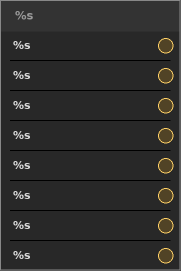
VISUALIZATION FRM_8BitPairDisplay  // 181x271
VAR_IN_OUT
    bBit0_1: BOOL;
    bBit1_1: BOOL;
    bBit2_1: BOOL;
    bBit3_1: BOOL;
    bBit4_1: BOOL;
    bBit5_1: BOOL;
    bBit6_1: BOOL;
    bBit7_1: BOOL;
    
    bBit0_2: BOOL;
    bBit1_2: BOOL;
    bBit2_2: BOOL;
    bBit3_2: BOOL;
    bBit4_2: BOOL;
    bBit5_2: BOOL;
    bBit6_2: BOOL;
    bBit7_2: BOOL;
END_VAR
VAR_INPUT
    sName: STRING;	

    sBitPair0: STRING;
    sBitPair1: STRING;
    sBitPair2: STRING;
    sBitPair3: STRING;
    sBitPair4: STRING;
    sBitPair5: STRING;
    sBitPair6: STRING;
    sBitPair7: STRING;	
END_VAR
    Rectangle (0,30 181x241)
    Textfield (10,40 141x11), "%s", text variable: sBitPair0
    Textfield (10,70 141x11), "%s", text variable: sBitPair1
    Textfield (10,100 141x11), "%s", text variable: sBitPair2
    Textfield (10,130 141x11), "%s", text variable: sBitPair3
    Textfield (10,160 141x11), "%s", text variable: sBitPair4
    Textfield (10,190 151x11), "%s", text variable: sBitPair5
    Textfield (10,220 141x11), "%s", text variable: sBitPair6
    Textfield (10,250 141x11), "%s", text variable: sBitPair7
    Line (10,60) (170,60)
    Line (10,90) (170,90)
    Line (10,120) (170,120)
    Line (10,150) (170,150)
    Line (10,180) (170,180)
    Line (10,210) (170,210)
    Line (10,240) (170,240)
    Textfield (0,0 181x31), "%s", text variable: sName
    Ellipse (158,38 15x15), colour toggle: bBit0_1 AND bBit0_2
    Ellipse (158,68 15x15), colour toggle: bBit1_1 AND bBit1_2
    Ellipse (158,98 15x15), colour toggle: bBit2_1 AND bBit2_2
    Ellipse (158,128 15x15), colour toggle: bBit3_1 AND bBit3_2
    Ellipse (158,158 15x15), colour toggle: bBit4_1 AND bBit4_2
    Ellipse (158,188 15x15), colour toggle: bBit5_1 AND bBit5_2
    Ellipse (158,218 15x15), colour toggle: bBit6_1 AND bBit6_2
    Ellipse (158,248 15x15), colour toggle: bBit7_1 AND bBit7_2
    Ellipse (158,38 15x15), invisible if: NOT (bBit0_1 XOR bBit0_2)
    Ellipse (158,68 15x15), invisible if: NOT (bBit1_1 XOR bBit1_2)
    Ellipse (158,98 15x15), invisible if: NOT (bBit2_1 XOR bBit2_2)
    Ellipse (158,128 15x15), invisible if: NOT (bBit3_1 XOR bBit3_2)
    Ellipse (158,158 15x15), invisible if: NOT (bBit4_1 XOR bBit4_2)
    Ellipse (158,188 15x15), invisible if: NOT (bBit5_1 XOR bBit5_2)
    Ellipse (158,218 15x15), invisible if: NOT (bBit6_1 XOR bBit6_2)
    Ellipse (158,248 15x15), invisible if: NOT (bBit7_1 XOR bBit7_2)
END_VISUALIZATION

(* stored: Version 1.1.0.1
   Visu FRM_8BitPairDisplay: Id {1f49f322-4436-0934-2d00-4a8ebd4d2a9b} *)
